Fanuc KAREL source: KA00097.KL

PROGRAM KA00097
%NOLOCKGROUP
VAR
  SRC: VECTOR
  DST: INTEGER
BEGIN
  SRC.X = 1.0
  DST = SRC
END KA00097
